(* IEC 61131-3 sources: llm-plc-st-eval/data/processed_definitivo/gpt-4o-2024-08-06/C7/zero_shot, 3 files *)

(* ---- ejec_1.st ---- *)
FUNCTION_BLOCK FB_Contador
VAR_INPUT
    sensorPieza : BOOL;   // Contacto normalmente abierto del sensor de pieza
    btnReset : BOOL;      // Contacto normalmente abierto para resetear el contador
END_VAR

VAR_OUTPUT
    loteListo : BOOL;     // Bobina que indica si el lote está listo
    cuenta : INT;         // Valor actual del contador
END_VAR

VAR
    C1 : CTU;             // Contador ascendente
END_VAR

// Inicialización del contador ascendente
C1(CU := sensorPieza, RESET := btnReset, PV := 12);

// Asignación de la salida del contador a la bobina loteListo
loteListo := C1.Q;

// Transferencia del valor actual del contador a la variable de salida cuenta
cuenta := C1.CV;
END_FUNCTION_BLOCK

(* ---- ejec_2.st ---- *)
FUNCTION_BLOCK FB_Contador
VAR_INPUT
    sensorPieza : BOOL;  // Contacto normalmente abierto para el sensor de pieza
    btnReset : BOOL;     // Contacto normalmente abierto para el botón de reset
END_VAR

VAR_OUTPUT
    loteListo : BOOL;    // Bobina que indica si el lote está listo
    cuenta : INT;        // Valor actual del contador
END_VAR

VAR
    C1 : CTU;            // Contador ascendente
END_VAR

// Inicialización del contador ascendente
C1(CU := sensorPieza, RESET := btnReset, PV := 12);

// Asignación de la salida del contador a la bobina loteListo
loteListo := C1.Q;

// Transferencia del valor actual del contador a la variable cuenta
cuenta := C1.CV;
END_FUNCTION_BLOCK

(* ---- ejec_3.st ---- *)
FUNCTION_BLOCK FB_Contador
VAR_INPUT
    sensorPieza : BOOL; // Contacto normalmente abierto para el sensor de pieza
    btnReset : BOOL;    // Contacto normalmente abierto para el botón de reset
END_VAR

VAR_OUTPUT
    loteListo : BOOL;   // Bobina que indica si el lote está listo
    cuenta : INT;       // Valor actual del contador
END_VAR

VAR
    C1 : CTU;           // Contador ascendente
END_VAR

// Configuración del contador ascendente
C1(CU := sensorPieza, RESET := btnReset, PV := 12);

// Asignación de la salida del contador a la bobina loteListo
loteListo := C1.Q;

// Transferencia del valor actual del contador a la variable cuenta
cuenta := C1.CV;
END_FUNCTION_BLOCK
